// TIA Portal V20 export
// export: Created 2026-10-19T18:37:18.2264528Z, ExportSetting WithDefaults, DisplayName Totally Integrated Automation Portal, DisplayVersion V20 Update 6, DisplayName TIA Portal Openness, DisplayVersion V20 Update 6, DisplayName TIA Portal Version Control Interface, DisplayVersion V20 Update 6, DisplayName SINAMICS Startdrive Advanced, DisplayVersion V20 SP1, DisplayName SINAMICS Startdrive G130, G150, S120, S150, SINAMICS MV, G220, S200, S210, DisplayVersion V20 SP1, DisplayName SINAMICS Startdrive G110M, G120, G120C, G120D, G120P, G115D, DisplayVersion V20 SP1, DisplayName STEP 7 Professional, DisplayVersion V20 Update 6, DisplayName STEP 7 Safety, DisplayVersion V20 Update 2, DisplayName WinCC Basic/Comfort/Advanced, DisplayVersion V20 Update 6, DisplayName WinCC Unified, DisplayVersion V20 Update 6
DATA_BLOCK "PopUp_Screens_1"   // DB51
{ S7_Optimized_Access := 'TRUE' }
VERSION : 0.1
// stored: AutoNumber true, DBAccessibleFromOPCUA true, IsOnlyStoredInLoadMemory false, IsRetainMemResEnabled false, IsWriteProtectedInAS false, MemoryReserve 100
   VAR
      LE_Speed : Array[1..6] of DInt;
      LE_Warnings : Array[1..6] of Byte;
      LE_Status : Array[1..6] of Bool;
      LE_Quality_Value : Array[1..6] of Int;
      LE_X_Unsafe_Position : Array[1..6] of UInt;
      LE_Quality_Decoded_Codes : Array[1..6] of UInt;
      LE_Bypass : Array[1..6] of DInt;
      AE_Speed : Array[1..6] of DInt;
      AE_Status_2 : Array[1..6] of UInt;
      AE_Control_Word_2 : Array[1..6] of UInt;
      AE_Position_1 : Array[1..6] of Bool;
      AE_Position_2 : Array[1..6] of Bool;
      AE_Status_1 : Array[1..6] of Bool;
      AE_Control_Word_1 : Array[1..6] of Bool;
      BCD_Disable_Trigger_HMI : Array[1..6] of Bool;
      BCD_Enable_Trigger_HMI : Array[1..6] of Bool;
      BCD_Error_HMI : Array[1..6] of Bool;
      BCD_Start_Comm_Test_HMI : Array[1..6] of Bool;
      BCD_Test_Ok_HMI : Array[1..6] of Bool;
      BCD_Execute_Function : Array[1..6] of Bool;
      BCD_RdDone : Array[1..6] of Bool;
      BCD_ReqDone : Array[1..6] of Bool;
      BCD_ReqBusy : Array[1..6] of Bool;
   END_VAR
BEGIN
END_DATA_BLOCK
